Fanuc KAREL source: KA00156.KL

PROGRAM KA00156
%NOLOCKGROUP
VAR
  SRC: ARRAY[4] OF REAL
  DST: ARRAY[4] OF BOOLEAN
BEGIN
  DST = SRC
END KA00156
